SYSTEM PID_Whiteboard (* Synthetic closed-loop example only; unmapped; native validation pending *)
  APPLICATION PID_Simulation
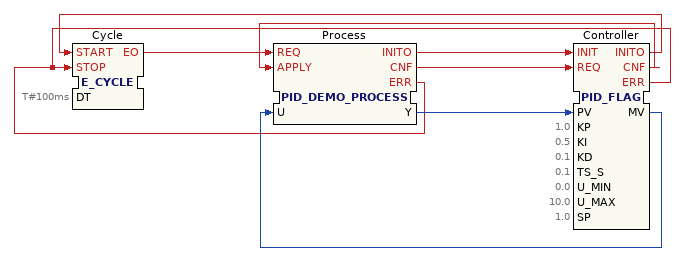
    FBS
      Cycle : E_CYCLE(DT := T#100ms);
      Process : PID_DEMO_PROCESS;
      Controller : PID_FLAG(KP := 1.0, KI := 0.5, KD := 0.1, TS_S := 0.1, U_MIN := 0.0, U_MAX := 10.0, SP := 1.0);
    END_FBS
    EVENT_CONNECTIONS
      Process.INITO TO Controller.INIT;
      Controller.INITO TO Cycle.START;
      Cycle.EO TO Process.REQ;
      Process.CNF TO Controller.REQ;
      Controller.CNF TO Process.APPLY;
      Process.ERR TO Cycle.STOP;
      Controller.ERR TO Cycle.STOP;
    END_CONNECTIONS
    DATA_CONNECTIONS
      Process.Y TO Controller.PV;
      Controller.MV TO Process.U;
    END_CONNECTIONS
  END_APPLICATION
  DEVICE LocalPID : FORTE_PC(MGR_ID := "localhost:61499")
    {SET_ATTRIBUTE(Profile, HOLOBLOC)} (* device profile *)
    RESOURCE EMB_RES : EMB_RES
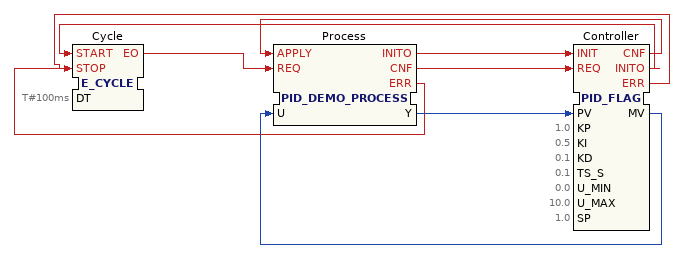
      FBS
        Controller : PID_FLAG(KP := 1.0, KI := 0.5, KD := 0.1, TS_S := 0.1, U_MIN := 0.0, U_MAX := 10.0, SP := 1.0);
        Process : PID_DEMO_PROCESS;
        Cycle : E_CYCLE(DT := T#100ms);
      END_FBS
      EVENT_CONNECTIONS
        Controller.CNF TO Process.APPLY;
        Process.INITO TO Controller.INIT;
        Process.CNF TO Controller.REQ;
        Controller.INITO TO Cycle.START;
        Process.ERR TO Cycle.STOP;
        Controller.ERR TO Cycle.STOP;
        Cycle.EO TO Process.REQ;
      END_CONNECTIONS
      DATA_CONNECTIONS
        Controller.MV TO Process.U;
        Process.Y TO Controller.PV;
      END_CONNECTIONS
    END_RESOURCE
  END_DEVICE
  MAPPINGS
    PID_Simulation.Controller ON LocalPID.EMB_RES.Controller;
    PID_Simulation.Process ON LocalPID.EMB_RES.Process;
    PID_Simulation.Cycle ON LocalPID.EMB_RES.Cycle;
  END_MAPPINGS
END_SYSTEM
